Fanuc KAREL source: ko00082.KL

-- PROVISIONAL review KL for V1013-1; original PC SHA256 0165b1b045f976cb1645a8493d0c2cb55e726082bba1fff14665324bfd7a1ecc
-- Incomplete behavior may be omitted. Consult companion uncertainty JSON. Do not deploy.
PROGRAM KO00082
%NOLOCKGROUP
BEGIN
  -- UNRESOLVED_PC offsets 5-12; opcodes 9D,23
  -- UNRESOLVED_PC offsets 17-66; opcodes 27,27,49,7E,AD,22,1C,22,31,7E,4A
  -- UNRESOLVED_PC offsets 71-75; opcodes 7F
END KO00082
